// TIA Portal project "000000000000-某某-自动配料模拟系统" (V15)

(* hardware
DEVICE "S7-1200 station_1"  S7-1200 Station
   slot 0: "Rack_0"  S7-1200 Rack  Rack  V1.0
   slot 1: "PLC_1"  CPU 1214C DC/DC/Rly  6ES7 214-1HG40-0XB0  V4.2
*)

// ===== PLC "PLC_1"  CPU 1214C DC/DC/Rly =====

VAR_GLOBAL   // PLC tag table "默认变量表"
   "System_Byte" AT %MB10 : Byte;
   "FirstScan" AT %M10.0 : Bool;
   "DiagStatusUpdate" AT %M10.1 : Bool;
   "AlwaysTRUE" AT %M10.2 : Bool;
   "AlwaysFALSE" AT %M10.3 : Bool;
   "M0.0" AT %M0.0 : Bool;
   "M0.1" AT %M0.1 : Bool;
   "M0.2" AT %M0.2 : Bool;
   "M0.3" AT %M0.3 : Bool;
   "M0.4" AT %M0.4 : Bool;
   "M0.5" AT %M0.5 : Bool;
   "M0.6" AT %M0.6 : Bool;
   "M0.7" AT %M0.7 : Bool;
   "M1.0" AT %M1.0 : Bool;
   "M1.1" AT %M1.1 : Bool;
   "M1.2" AT %M1.2 : Bool;
   "M1.3" AT %M1.3 : Bool;
   "M1.4" AT %M1.4 : Bool;
   "M1.5" AT %M1.5 : Bool;
   "M1.6" AT %M1.6 : Bool;
   "启动" AT %I0.0 : Bool;
   "停止" AT %I0.1 : Bool;
   "物料传感器" AT %I0.2 : Bool;
   "限位开关1" AT %I0.3 : Bool;
   "限位开关2" AT %I0.4 : Bool;
   "出料阀" AT %Q0.0 : Bool;
   "进料阀" AT %Q0.1 : Bool;
   "L1" AT %Q0.2 : Bool;
   "L2" AT %Q0.3 : Bool;
   "KM1" AT %Q1.0 : Bool;
   "KM2" AT %Q1.1 : Bool;
   "KM3" AT %Q1.2 : Bool;
   "KM4" AT %Q1.3 : Bool;
   "Tag_1" AT %MD10 : Time;
   "Tag_2" AT %MD14 : Time;
   "Tag_3" AT %MD18 : Time;
   "Tag_4" AT %MD22 : Time;
   "Tag_5" AT %MD26 : Time;
   "Tag_6" AT %MD30 : Time;
   "Tag_7" AT %MD34 : Time;
   "Tag_8" AT %MD38 : Time;
   "Tag_9" AT %MD42 : Time;
END_VAR

// folder: System blocks/Program resources

DATA_BLOCK "T1"   // DB1
{ S7_Optimized_Access := 'TRUE' }
AUTHOR : Simatic
FAMILY : IEC
NAME : IEC_TMR
VERSION : 1.0
// stored: InstanceOfName IEC_TIMER
"IEC_TIMER"
BEGIN
END_DATA_BLOCK

DATA_BLOCK "T2"   // DB2
{ S7_Optimized_Access := 'TRUE' }
AUTHOR : Simatic
FAMILY : IEC
NAME : IEC_TMR
VERSION : 1.0
// stored: InstanceOfName IEC_TIMER
"IEC_TIMER"
BEGIN
END_DATA_BLOCK

DATA_BLOCK "T3"   // DB3
{ S7_Optimized_Access := 'TRUE' }
AUTHOR : Simatic
FAMILY : IEC
NAME : IEC_TMR
VERSION : 1.0
// stored: InstanceOfName IEC_TIMER
"IEC_TIMER"
BEGIN
END_DATA_BLOCK

DATA_BLOCK "T4"   // DB4
{ S7_Optimized_Access := 'TRUE' }
AUTHOR : Simatic
FAMILY : IEC
NAME : IEC_TMR
VERSION : 1.0
// stored: InstanceOfName IEC_TIMER
"IEC_TIMER"
BEGIN
END_DATA_BLOCK

DATA_BLOCK "T5"   // DB5
{ S7_Optimized_Access := 'TRUE' }
AUTHOR : Simatic
FAMILY : IEC
NAME : IEC_TMR
VERSION : 1.0
// stored: InstanceOfName IEC_TIMER
"IEC_TIMER"
BEGIN
END_DATA_BLOCK

DATA_BLOCK "T6"   // DB6
{ S7_Optimized_Access := 'TRUE' }
AUTHOR : Simatic
FAMILY : IEC
NAME : IEC_TMR
VERSION : 1.0
// stored: InstanceOfName IEC_TIMER
"IEC_TIMER"
BEGIN
END_DATA_BLOCK

DATA_BLOCK "T7"   // DB7
{ S7_Optimized_Access := 'TRUE' }
AUTHOR : Simatic
FAMILY : IEC
NAME : IEC_TMR
VERSION : 1.0
// stored: InstanceOfName IEC_TIMER
"IEC_TIMER"
BEGIN
END_DATA_BLOCK

DATA_BLOCK "T8"   // DB8
{ S7_Optimized_Access := 'TRUE' }
AUTHOR : Simatic
FAMILY : IEC
NAME : IEC_TMR
VERSION : 1.0
// stored: InstanceOfName IEC_TIMER
"IEC_TIMER"
BEGIN
END_DATA_BLOCK

DATA_BLOCK "保护"   // DB9
{ S7_Optimized_Access := 'TRUE' }
AUTHOR : Simatic
FAMILY : IEC
NAME : IEC_TMR
VERSION : 1.0
// stored: InstanceOfName IEC_TIMER
"IEC_TIMER"
BEGIN
END_DATA_BLOCK

// folder: (top level)

ORGANIZATION_BLOCK "Main"   // OB1, LAD, ProgramCycle
TITLE = "Main Program Sweep (Cycle)"
{ S7_Optimized_Access := 'TRUE' }
VERSION : 0.1
   VAR_INPUT
      Initial_Call : Bool;   // Initial call of this OB
      Remanence : Bool;   // =True, if remanent data are available
   END_VAR
   VAR_TEMP   // added for the SCL form of the ladder/FBD networks
      _w1 : Bool;
      _w2 : Bool;
      _w3 : Bool;
      _w4 : Bool;
      _w5 : Bool;
      _w6 : Bool;
      _w7 : Bool;
      _w8 : Bool;
   END_VAR
BEGIN

REGION Network 1
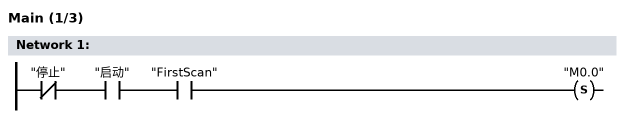
   RUNG wire#powerrail
      I_Contact( "停止" )
      Contact( "启动" )
      Contact( "FirstScan" )
      S_Coil( "M0.0" )
   END_RUNG
   // the same network as SCL:
   IF NOT "停止" AND "启动" AND "FirstScan" THEN "M0.0" := TRUE; END_IF;
END_REGION

REGION Network 2
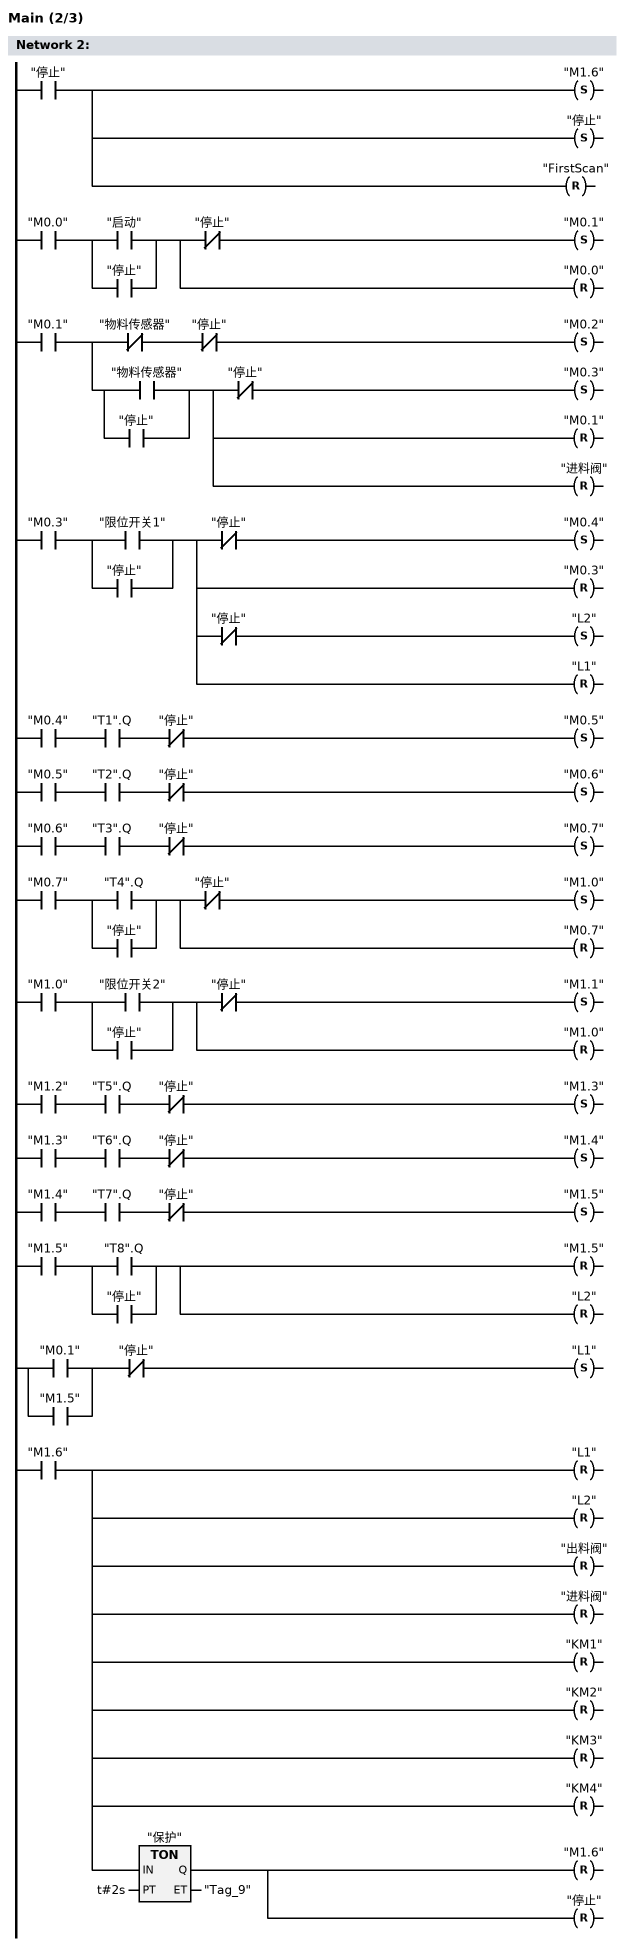
   IF "停止" THEN "M1.6" := TRUE; END_IF;
   #_w1 := "停止";
   IF #_w1 THEN
       "停止" := TRUE;
       "FirstScan" := FALSE;
   END_IF;
   #_w2 := "M0.0" AND ("启动" OR "停止");
   IF #_w2 AND NOT "停止" THEN "M0.1" := TRUE; END_IF;
   IF #_w2 THEN "M0.0" := FALSE; END_IF;
   IF "M0.1" AND NOT "物料传感器" AND NOT "停止" THEN "M0.2" := TRUE; END_IF;
   #_w3 := "M0.1" AND ("物料传感器" OR "停止");
   IF #_w3 AND NOT "停止" THEN "M0.3" := TRUE; END_IF;
   IF #_w3 THEN
       "M0.1" := FALSE;
       "进料阀" := FALSE;
   END_IF;
   #_w4 := "M0.3" AND ("限位开关1" OR "停止");
   IF #_w4 AND NOT "停止" THEN "M0.4" := TRUE; END_IF;
   IF #_w4 THEN "M0.3" := FALSE; END_IF;
   IF #_w4 AND NOT "停止" THEN "L2" := TRUE; END_IF;
   IF #_w4 THEN "L1" := FALSE; END_IF;
   IF "M0.4" AND "T1".Q AND NOT "停止" THEN "M0.5" := TRUE; END_IF;
   IF "M0.5" AND "T2".Q AND NOT "停止" THEN "M0.6" := TRUE; END_IF;
   IF "M0.6" AND "T3".Q AND NOT "停止" THEN "M0.7" := TRUE; END_IF;
   #_w5 := "M0.7" AND ("T4".Q OR "停止");
   IF #_w5 AND NOT "停止" THEN "M1.0" := TRUE; END_IF;
   IF #_w5 THEN "M0.7" := FALSE; END_IF;
   #_w6 := "M1.0" AND ("限位开关2" OR "停止");
   IF #_w6 AND NOT "停止" THEN "M1.1" := TRUE; END_IF;
   IF #_w6 THEN "M1.0" := FALSE; END_IF;
   IF "M1.2" AND "T5".Q AND NOT "停止" THEN "M1.3" := TRUE; END_IF;
   IF "M1.3" AND "T6".Q AND NOT "停止" THEN "M1.4" := TRUE; END_IF;
   IF "M1.4" AND "T7".Q AND NOT "停止" THEN "M1.5" := TRUE; END_IF;
   #_w7 := "M1.5" AND ("T8".Q OR "停止");
   IF #_w7 THEN
       "M1.5" := FALSE;
       "L2" := FALSE;
   END_IF;
   IF ("M0.1" OR "M1.5") AND NOT "停止" THEN "L1" := TRUE; END_IF;
   IF "M1.6" THEN
       "L1" := FALSE;
       "L2" := FALSE;
       "出料阀" := FALSE;
       "进料阀" := FALSE;
       "KM1" := FALSE;
       "KM2" := FALSE;
       "KM3" := FALSE;
       "KM4" := FALSE;
   END_IF;
   "保护".TON(IN := "M1.6", PT := t#2s, ET => "Tag_9");
   IF "保护".Q THEN
       "M1.6" := FALSE;
       "停止" := FALSE;
   END_IF;
END_REGION

REGION Network 3
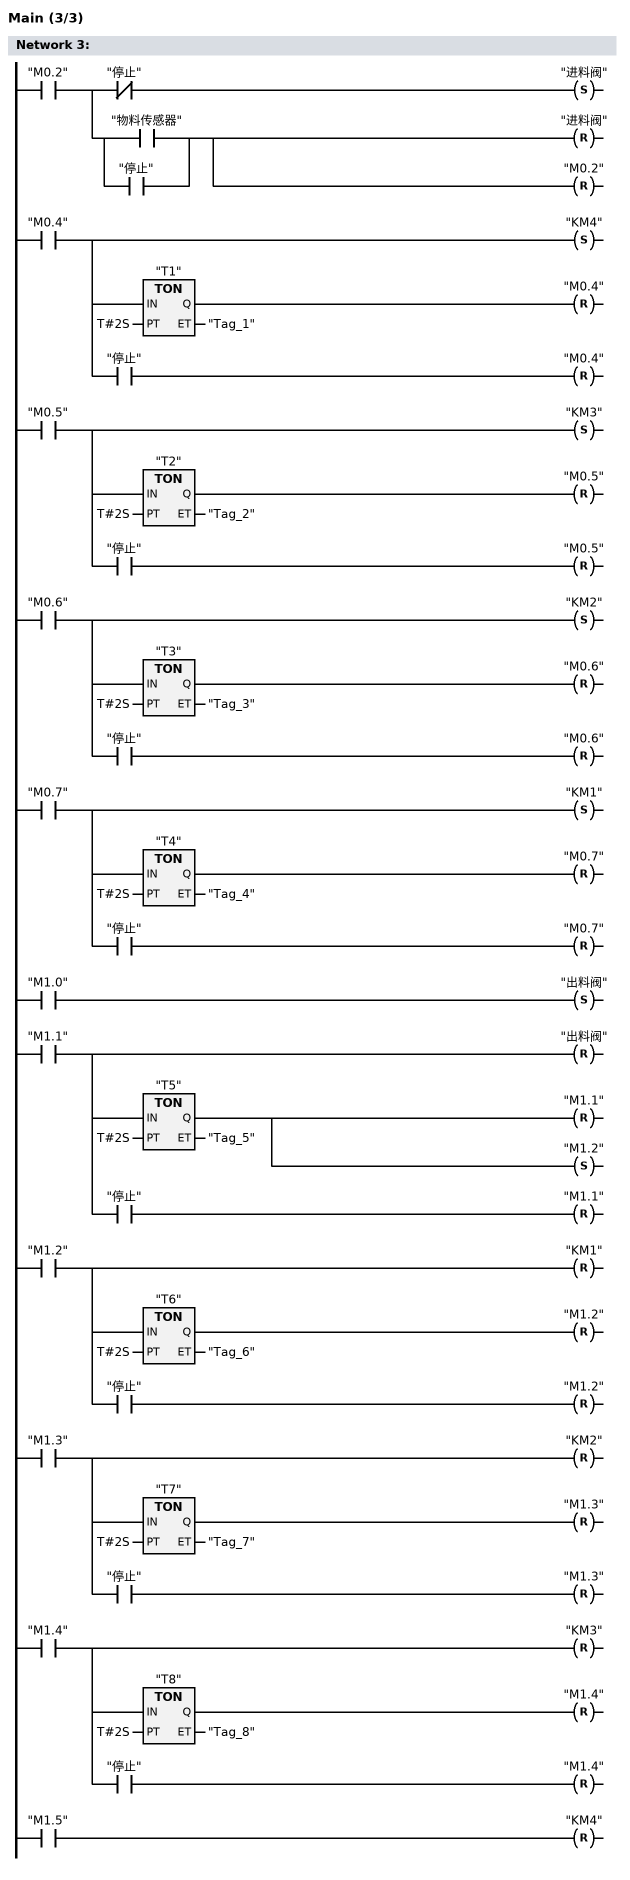
   IF "M0.2" AND NOT "停止" THEN "进料阀" := TRUE; END_IF;
   IF "M0.2" AND ("物料传感器" OR "停止") THEN
       "进料阀" := FALSE;
       "M0.2" := FALSE;
   END_IF;
   IF "M0.4" THEN "KM4" := TRUE; END_IF;
   "T1".TON(IN := "M0.4", PT := T#2S, ET => "Tag_1");
   #_w1 := "M0.4";
   IF "T1".Q THEN "M0.4" := FALSE; END_IF;
   IF #_w1 AND "停止" THEN "M0.4" := FALSE; END_IF;
   IF "M0.5" THEN "KM3" := TRUE; END_IF;
   "T2".TON(IN := "M0.5", PT := T#2S, ET => "Tag_2");
   #_w2 := "M0.5";
   IF "T2".Q THEN "M0.5" := FALSE; END_IF;
   IF #_w2 AND "停止" THEN "M0.5" := FALSE; END_IF;
   IF "M0.6" THEN "KM2" := TRUE; END_IF;
   "T3".TON(IN := "M0.6", PT := T#2S, ET => "Tag_3");
   #_w3 := "M0.6";
   IF "T3".Q THEN "M0.6" := FALSE; END_IF;
   IF #_w3 AND "停止" THEN "M0.6" := FALSE; END_IF;
   IF "M0.7" THEN "KM1" := TRUE; END_IF;
   "T4".TON(IN := "M0.7", PT := T#2S, ET => "Tag_4");
   #_w4 := "M0.7";
   IF "T4".Q THEN "M0.7" := FALSE; END_IF;
   IF #_w4 AND "停止" THEN "M0.7" := FALSE; END_IF;
   IF "M1.0" THEN "出料阀" := TRUE; END_IF;
   IF "M1.1" THEN "出料阀" := FALSE; END_IF;
   "T5".TON(IN := "M1.1", PT := T#2S, ET => "Tag_5");
   #_w5 := "M1.1";
   IF "T5".Q THEN
       "M1.1" := FALSE;
       "M1.2" := TRUE;
   END_IF;
   IF #_w5 AND "停止" THEN "M1.1" := FALSE; END_IF;
   IF "M1.2" THEN "KM1" := FALSE; END_IF;
   "T6".TON(IN := "M1.2", PT := T#2S, ET => "Tag_6");
   #_w6 := "M1.2";
   IF "T6".Q THEN "M1.2" := FALSE; END_IF;
   IF #_w6 AND "停止" THEN "M1.2" := FALSE; END_IF;
   IF "M1.3" THEN "KM2" := FALSE; END_IF;
   "T7".TON(IN := "M1.3", PT := T#2S, ET => "Tag_7");
   #_w7 := "M1.3";
   IF "T7".Q THEN "M1.3" := FALSE; END_IF;
   IF #_w7 AND "停止" THEN "M1.3" := FALSE; END_IF;
   IF "M1.4" THEN "KM3" := FALSE; END_IF;
   "T8".TON(IN := "M1.4", PT := T#2S, ET => "Tag_8");
   #_w8 := "M1.4";
   IF "T8".Q THEN "M1.4" := FALSE; END_IF;
   IF #_w8 AND "停止" THEN "M1.4" := FALSE; END_IF;
   IF "M1.5" THEN "KM4" := FALSE; END_IF;
END_REGION
END_ORGANIZATION_BLOCK